Staubli VAL3: getProgItemIndex.pgx

public program getProgItemIndex(string x_sKey, string x_sSelProgItem, num& x_nIndex)
  local num l_nSize
  local bool l_bResult
begin
  call getProgItemSize(x_sKey,l_nSize)
  if l_nSize==1 and progTemp:pProgItem[x_sKey].pProgTemplate[0].sTRAJname==""
    x_nIndex=0
  else
    toNum(x_sSelProgItem,x_nIndex,l_bResult)
  endIf

end
